(* IEC 61131-3 sources: 2026_Projet_YGO_ExcavatriceDragage/CODE/DIAG, 4 files *)

(* ---- E_DiagState.st ---- *)
(* ═══════════════════════════════════════════════════════════════
   🚦 E_DiagState — Énumération des phases de diagnostic bus
   ═══════════════════════════════════════════════════════════════ *)
TYPE E_DiagState :
(
    DISABLED   := 0,  (* Désactivé (surveillance non active) *)
    READY      := 1,  (* Prêt (opérationnel, pas de défaut) *)
    INIT       := 2,  (* Initialisation en cours / Recherche de réseau *)
    MONITORING := 3,  (* Surveillance active (états transitoires) *)
    ERROR      := 4   (* Présence anomalie de communication *)
);
END_TYPE

(* ---- ST_DeviceDiag.st ---- *)
(* ═══════════════════════════════════════════════════════════════
   📡 ST_DeviceDiag — Structure diagnostic d'un esclave ou bus
   ═══════════════════════════════════════════════════════════════ *)
TYPE ST_DeviceDiag :
STRUCT
    Online         : BOOL;        (* Esclave visible sur le bus *)
    Operational    : BOOL;        (* Esclave en mode OP (opérationnel) *)
    Error          : BOOL;        (* Signal de défaut actif pour cet esclave *)
    ErrorId        : WORD;        (* Code défaut détaillé *)
    State          : E_DiagState; (* Phase courante du cycle de diagnostic *)
    StateAtError   : E_DiagState; (* Instantané de la phase lors de l'anomalie *)
END_STRUCT
END_TYPE

(* ---- FB_DiagCanOpen.st ---- *)
(* ═══════════════════════════════════════════════════════════════
   📡 FB_DiagCanOpen — Diagnostic de communication bus CANopen / Joystick
   ═══════════════════════════════════════════════════════════════ *)
FUNCTION_BLOCK PUBLIC FB_DiagCanOpen
VAR_INPUT
    Enable          : BOOL;        (* Active la surveillance CAN *)
    Reset           : BOOL;        (* Front d'acquittement des défauts *)
    CanOnline       : BOOL;        (* Trame joystick reçue (TRUE = OK) *)
    CanOperational  : BOOL;        (* Joystick en mode opérationnel (TRUE = OK) *)
END_VAR
VAR_OUTPUT
    Ready           : BOOL;        (* Logique de surveillance active *)
    Busy            : BOOL;        (* Non utilisé (conformité interface) *)
    Done            : BOOL;        (* Non utilisé *)
    Error           : BOOL;        (* Présence anomalie de communication *)
    ErrorId         : WORD;        (* Code défaut global résumé *)
    State           : E_DiagState; (* Phase courante du cycle de diag *)
    StateAtError    : E_DiagState; (* Phase figée à l'apparition de l'erreur *)
    busCanOpen      : ST_DeviceDiag;  (* Diagnostics bus CANopen *)
    Joystick        : ST_DeviceDiag;  (* Diagnostics esclave Joystick *)
END_VAR
VAR
    ResetEdge       : R_TRIG;      (* Détecteur front de reset *)
END_VAR

// 🛑 1. GATE : Désactivation logique si Enable = FALSE
IF NOT Enable THEN
    Ready := FALSE;
    State := E_DiagState.DISABLED;
    Joystick.State := E_DiagState.DISABLED;
    Joystick.Online := FALSE;
    Joystick.Operational := FALSE;
    Joystick.Error := FALSE;
    Joystick.ErrorId := 16#0000;
    Error := FALSE;
    ErrorId := 16#0000;
    RETURN;
END_IF;

Ready := TRUE;

// 🔑 2. RESET FRONT — Efface les défauts si la cause a disparu
ResetEdge(CLK := Reset);
IF ResetEdge.Q THEN
    IF (CanOnline AND CanOperational) THEN
        Joystick.ErrorId := 16#0000;
        StateAtError := E_DiagState.DISABLED;
    END_IF;
END_IF;

// 🔍 3. DIAGNOSTIC JOYSTICK
// Bit 0 : Perte de communication CAN
IF NOT CanOnline THEN
    Joystick.ErrorId := 16#0001;  (* Perte liaison CAN joystick *)
    Joystick.Online := FALSE;
ELSE
    Joystick.Online := TRUE;
    IF ResetEdge.Q THEN
        Joystick.ErrorId := Joystick.ErrorId AND 16#FFFE;
    END_IF;
END_IF;

// Bit 1 : Mode non-opérationnel (esclave CANopen en pré-op ou défaut)
IF NOT CanOperational THEN
    Joystick.ErrorId := Joystick.ErrorId OR 16#0002;  (* Joystick pas opérationnel *)
    Joystick.Operational := FALSE;
ELSE
    Joystick.Operational := TRUE;
    IF ResetEdge.Q THEN
        Joystick.ErrorId := Joystick.ErrorId AND 16#FFFD;
    END_IF;
END_IF;

// 🚦 4. MACHINE D'ÉTAT JOYSTICK
IF Joystick.ErrorId <> 0 THEN
    Joystick.State := E_DiagState.ERROR;
    IF StateAtError = E_DiagState.DISABLED THEN
        StateAtError := State;
    END_IF;
ELSIF NOT (Joystick.Online AND Joystick.Operational) THEN
    Joystick.State := E_DiagState.INIT;
else
    Joystick.State := E_DiagState.READY;
END_IF;

State := Joystick.State;

// 📤 5. SORTIES GLOBALES
Joystick.Error := (Joystick.ErrorId <> 0);
Error := Joystick.Error;
ErrorId := Joystick.ErrorId;

busCanOpen.Operational := CanOnline;
busCanOpen.Online := CanOnline;

// Briques génériques pour conformité standard
Busy := FALSE;
Done := FALSE;

(* ---- FB_DiagEthercat.st ---- *)
(* ═══════════════════════════════════════════════════════════════
   📡 FB_DiagEthercat — Diagnostic de communication bus EtherCAT (3 esclaves)
   ═══════════════════════════════════════════════════════════════ *)
FUNCTION_BLOCK PUBLIC FB_DiagEthercat
VAR_INPUT
    Enable              : BOOL;        (* Active la surveillance EtherCAT *)
    Reset               : BOOL;        (* Front d'acquittement des défauts *)

    (* Variateur M3 (AC600_ECAT_Drive) *)
    VariateurWcState    : BOOL;        (* Working Counter variateur (FALSE = OK) *)
    VariateurSlaveState : WORD;        (* État esclave variateur (8 = OP) *)

    (* Encodeur M1 (COD1_CODEUR) *)
    EncoderM1WcState    : BOOL;        (* Working Counter M1 (FALSE = OK) *)
    EncoderM1SlaveState : WORD;        (* État esclave M1 (8 = OP) *)

    (* Encodeur M2 (COD2_CODEUR) *)
    EncoderM2WcState    : BOOL;        (* Working Counter M2 (FALSE = OK) *)
    EncoderM2SlaveState : WORD;        (* État esclave M2 (8 = OP) *)
END_VAR
VAR_OUTPUT
    Ready               : BOOL;        (* Logique de surveillance active *)
    Busy                : BOOL;        (* Non utilisé (conformité) *)
    Done                : BOOL;        (* Non utilisé *)
    Error               : BOOL;        (* Résumé anomalie de communication bus *)
    ErrorId             : WORD;        (* Code défaut global résumé *)
    State               : E_DiagState; (* Phase courante du diagnostic global *)
    StateAtError        : E_DiagState; (* Phase figée à l'apparition de l'erreur *)
    BusEthercat         : ST_DeviceDiag;  (* Diagnostics bus EtherCAT *)
    Variateur           : ST_DeviceDiag;  (* Diagnostics esclave AC600 *)
    EncoderM1           : ST_DeviceDiag;  (* Diagnostics esclave COD1 *)
    EncoderM2           : ST_DeviceDiag;  (* Diagnostics esclave COD2 *)
END_VAR
VAR
    ResetEdge           : R_TRIG;      (* Détecteur front de reset *)
END_VAR

// 🛑 1. GATE : Désactivation si Enable = FALSE
IF NOT Enable THEN
    Ready := FALSE;
    State := E_DiagState.DISABLED;
    Variateur.State := E_DiagState.DISABLED;
    EncoderM1.State := E_DiagState.DISABLED;
    EncoderM2.State := E_DiagState.DISABLED;
    Variateur.Online := FALSE;
    EncoderM1.Online := FALSE;
    EncoderM2.Online := FALSE;
    Variateur.Operational := FALSE;
    EncoderM1.Operational := FALSE;
    EncoderM2.Operational := FALSE;
    Variateur.Error := FALSE;
    EncoderM1.Error := FALSE;
    EncoderM2.Error := FALSE;
    Error := FALSE;
    ErrorId := 16#0000;
    RETURN;
END_IF;

Ready := TRUE;

// 🔑 2. RESET FRONT
ResetEdge(CLK := Reset);

// 🔍 3. DIAGNOSTIC VARIATEUR (AC600_ECAT_Drive / Translation M3)
Variateur.Online := NOT VariateurWcState;
Variateur.Operational := Variateur.Online AND (VariateurSlaveState = 8);

IF NOT Variateur.Online THEN
    Variateur.ErrorId := 16#0010;  (* Perte liaison physique variateur *)
ELSE
    IF ResetEdge.Q THEN
        Variateur.ErrorId := Variateur.ErrorId AND 16#FFEF;
    END_IF;
END_IF;

IF NOT Variateur.Operational AND Variateur.Online THEN
    Variateur.ErrorId := Variateur.ErrorId OR 16#0011;  (* Variateur pré-opérationnel *)
ELSE
    IF ResetEdge.Q THEN
        Variateur.ErrorId := Variateur.ErrorId AND 16#FFEE;
    END_IF;
END_IF;

// 🔍 4. DIAGNOSTIC ENCODEUR M1 (COD1_CODEUR / WinchM1)
EncoderM1.Online := NOT EncoderM1WcState;
EncoderM1.Operational := EncoderM1.Online AND (EncoderM1SlaveState = 8);

IF NOT EncoderM1.Online THEN
    EncoderM1.ErrorId := 16#0020;  (* Perte liaison encodeur M1 *)
ELSE
    IF ResetEdge.Q THEN
        EncoderM1.ErrorId := EncoderM1.ErrorId AND 16#FFDF;
    END_IF;
END_IF;

IF NOT EncoderM1.Operational AND EncoderM1.Online THEN
    EncoderM1.ErrorId := EncoderM1.ErrorId OR 16#0021;  (* Encodeur M1 pré-opérationnel *)
ELSE
    IF ResetEdge.Q THEN
        EncoderM1.ErrorId := EncoderM1.ErrorId AND 16#FFDE;
    END_IF;
END_IF;

// 🔍 5. DIAGNOSTIC ENCODEUR M2 (COD2_CODEUR / WinchM2)
EncoderM2.Online := NOT EncoderM2WcState;
EncoderM2.Operational := EncoderM2.Online AND (EncoderM2SlaveState = 8);

IF NOT EncoderM2.Online THEN
    EncoderM2.ErrorId := 16#0030;  (* Perte liaison encodeur M2 *)
ELSE
    IF ResetEdge.Q THEN
        EncoderM2.ErrorId := EncoderM2.ErrorId AND 16#FFCF;
    END_IF;
END_IF;

IF NOT EncoderM2.Operational AND EncoderM2.Online THEN
    EncoderM2.ErrorId := EncoderM2.ErrorId OR 16#0031;  (* Encodeur M2 pré-opérationnel *)
ELSE
    IF ResetEdge.Q THEN
        EncoderM2.ErrorId := EncoderM2.ErrorId AND 16#FFCE;
    END_IF;
END_IF;

// 🚦 6. STATE MACHINES DE CHAQUE APPAREIL
IF Variateur.ErrorId <> 0 THEN
    Variateur.State := E_DiagState.ERROR;
ELSIF NOT Variateur.Online THEN
    Variateur.State := E_DiagState.INIT;
ELSIF Variateur.Operational THEN
    Variateur.State := E_DiagState.READY;
ELSE
    Variateur.State := E_DiagState.MONITORING;
END_IF;

IF EncoderM1.ErrorId <> 0 THEN
    EncoderM1.State := E_DiagState.ERROR;
ELSIF NOT EncoderM1.Online THEN
    EncoderM1.State := E_DiagState.INIT;
ELSIF EncoderM1.Operational THEN
    EncoderM1.State := E_DiagState.READY;
ELSE
    EncoderM1.State := E_DiagState.MONITORING;
END_IF;

IF EncoderM2.ErrorId <> 0 THEN
    EncoderM2.State := E_DiagState.ERROR;
ELSIF NOT EncoderM2.Online THEN
    EncoderM2.State := E_DiagState.INIT;
ELSIF EncoderM2.Operational THEN
    EncoderM2.State := E_DiagState.READY;
ELSE
    EncoderM2.State := E_DiagState.MONITORING;
END_IF;

// Fige la phase du diagnostic global sur le premier défaut
IF (Variateur.ErrorId <> 0 OR EncoderM1.ErrorId <> 0 OR EncoderM2.ErrorId <> 0) THEN
    IF StateAtError = E_DiagState.DISABLED THEN
        StateAtError := State;
    END_IF;
END_IF;

// 📤 7. RÉSUMÉ ET DÉFAUTS
Variateur.Error := (Variateur.ErrorId <> 0);
EncoderM1.Error := (EncoderM1.ErrorId <> 0);
EncoderM2.Error := (EncoderM2.ErrorId <> 0);

Error := (Variateur.Error OR EncoderM1.Error OR EncoderM2.Error);

ErrorId := 16#0000;
IF Variateur.Error THEN
    ErrorId := ErrorId OR 16#00F0;
END_IF;
IF EncoderM1.Error THEN
    ErrorId := ErrorId OR 16#0F00;
END_IF;
IF EncoderM2.Error THEN
    ErrorId := ErrorId OR 16#F000;
END_IF;

IF Error THEN
    State := E_DiagState.ERROR;
ELSIF NOT (Variateur.Operational AND EncoderM1.Operational AND EncoderM2.Operational) THEN
    State := E_DiagState.MONITORING;
ELSE
    State := E_DiagState.READY;
END_IF;

BusEthercat.Online := Variateur.Online AND EncoderM1.Online AND EncoderM2.Online;
BusEthercat.Operational := Variateur.Operational AND EncoderM1.Operational AND EncoderM2.Operational;

Busy := FALSE;
Done := FALSE;
